(* PLC project Vn_or2, Beckhoff Automation GmbH TwinCAT PLC Control 3.5.13.21 *)
(* stored: creationDateTime 1970-01-01T00:00:00 *)

PROGRAM Vn_or2

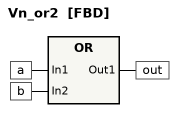
(* FBD diagram, written out as Structured Text *)
out := a OR b;
END_PROGRAM
